// TIA Portal V19 export
TYPE "ST_RECIPE"
   STRUCT
      Id : Int;
      "Name" : String;
      ProductName : String;
      Columns : Int;
      Rows : Int;
      ProductHeight : Int;
      Pattern1 : Bool;
      Pattern2 : Bool;
   END_STRUCT;
END_TYPE
